{attribute 'linkalways'} 
{attribute 'no_explicit_call' := 'This FB is a CLASS and must be accessed using methods or properties'}
{attribute 'enable_dynamic_creation'}
FUNCTION_BLOCK _ETcVnEdgeDetectionAlgorithm EXTENDS EnumDatatypeBase
VAR
	localData : ETcVnEdgeDetectionAlgorithm;
	activeData : REFERENCE TO ETcVnEdgeDetectionAlgorithm;
	enumBaseDatatype : _DINT(localData);
END_VAR

METHOD PRIVATE AddLocalEnumeration
VAR_INPUT
	Enumeration : T_MAXSTRING;
	Value : ETcVnEdgeDetectionAlgorithm;
END_VAR
AddEnumeration(Enumeration, Value);
END_METHOD

PROPERTY PUBLIC Address : PVOID
GET
Address := ADR(activeData);
END_GET
END_PROPERTY

METHOD PUBLIC ClearReference
VAR_INPUT
END_VAR
activeData REF= localData;
SetBaseDatatypeReference();
END_METHOD

METHOD PUBLIC Clone : I_Datatype
VAR
    pClone : POINTER TO _ETcVnEdgeDetectionAlgorithm;
END_VAR
pClone := __NEW(_ETcVnEdgeDetectionAlgorithm(InitialValue := Value));
Clone := pClone^;
END_METHOD

METHOD FB_init : BOOL
VAR_INPUT
	bInitRetains : BOOL; // if TRUE, the retain variables are initialized (warm start / cold start)
	bInCopyCode : BOOL;  // if TRUE, the instance afterwards gets moved into the copy code (online change)
	InitialValue : ETcVnEdgeDetectionAlgorithm;
END_VAR
localData := InitialValue;
AddBaseDatatype(enumBaseDatatype);
ClearReference();

AddLocalEnumeration('TCVN_EDA_INTERPOLATION', ETcVnEdgeDetectionAlgorithm.TCVN_EDA_INTERPOLATION);
AddLocalEnumeration('TCVN_EDA_APPROX_ERF', ETcVnEdgeDetectionAlgorithm.TCVN_EDA_APPROX_ERF);
AddLocalEnumeration('TCVN_EDA_APPROX_GAUSSIAN', ETcVnEdgeDetectionAlgorithm.TCVN_EDA_APPROX_GAUSSIAN);
END_METHOD

PROPERTY PUBLIC Identifier : T_MAXSTRING
GET
Identifier := 'ETcVnEdgeDetectionAlgorithm';
END_GET
END_PROPERTY

METHOD IsEnumeratorValueEqual : BOOL
VAR_INPUT
	Enumerator : I_KeyValueForwardEnumerator;
END_VAR
VAR
	storedValue : ETcVnEdgeDetectionAlgorithm;
END_VAR
IF NOT Enumerator.TryGet(storedValue) THEN
	RETURN;
END_IF

IsEnumeratorValueEqual := storedValue = activeData;
END_METHOD

METHOD PUBLIC MakeReferenceTo
VAR_INPUT
	ReferenceTarget : REFERENCE TO ETcVnEdgeDetectionAlgorithm;
END_VAR
activeData REF= ReferenceTarget;
SetBaseDatatypeReference();
END_METHOD

METHOD PROTECTED SetBaseDatatypeReference
VAR_INPUT
END_VAR
enumBaseDatatype.MakeReferenceTo(activeData);
END_METHOD

PROPERTY PUBLIC Size : UDINT
GET
Size := SIZEOF(activeData);
END_GET
END_PROPERTY

METHOD TryMakeReferenceTo : BOOL
VAR_INPUT
	Target : I_Datatype;
END_VAR
VAR
	pTargetData : POINTER TO ETcVnEdgeDetectionAlgorithm;
END_VAR
IF NOT IsEquivalentTo(Target) THEN
	RETURN;
END_IF

pTargetData := Target.Address;
activeData REF= pTargetData^;
SetBaseDatatypeReference();
TryMakeReferenceTo := TRUE;
END_METHOD

PROPERTY PUBLIC Value : ETcVnEdgeDetectionAlgorithm
GET
Value := activeData;
END_GET
SET
activeData := Value;
END_SET
END_PROPERTY

END_FUNCTION_BLOCK

(* stored: Version 1.1.0.1, ProductVersion 3.1.4024.13
   POU _ETcVnEdgeDetectionAlgorithm: Id {de3327d9-628b-0db8-070f-b6ec3e9cfed8}, SpecialFunc None
   Folder Core: Id {e035bb8f-f195-0321-2564-328d1d9e6354}
   Folder Protected: Id {24d363fe-2ee2-017f-0644-1bdf48376c97}
   Folder Customize: Id {5e2cb9a4-28a6-0918-2e91-0ebe8bb50e53}
   Folder Constructor: Id {163cf6a0-f511-071e-20fa-813a2df9bf96}
   Folder Private: Id {fa96855c-e46a-09e8-18d9-cd7d699408c7}
   Folder Protected: Id {81f72d85-df5c-0d10-25bf-c5676d71d58f}
   Method AddLocalEnumeration: Id {c7807dc8-fcd2-0167-2c69-db3e14617561}
   Property Address: Id {1c4d0320-6103-0427-3c85-658858caa5d9}
   Get Get: Id {2ceb24b0-bddc-0b13-0661-3c4ac1ff7d2a}
   Method ClearReference: Id {06331ef3-70e5-04b8-06bb-a3e7476cd189}
   Method Clone: Id {93dcc90a-ca49-0669-2de3-8775364a3c48}
   Method FB_init: Id {499c5acc-ee1f-048c-274d-37da243b2af5}
   Property Identifier: Id {73c0b194-9924-0dcf-2ac0-b517abdb4f5b}
   Get Get: Id {2391be6c-42a0-0570-0938-859bb6badf5f}
   Method IsEnumeratorValueEqual: Id {15a04b32-a76a-0a9a-0ce5-ab7589c338e2}
   Method MakeReferenceTo: Id {96185666-00ce-04b4-2ca1-41455ce3c251}
   Method SetBaseDatatypeReference: Id {9d4bfa6b-0ad5-0f35-2704-873b62a7c773}
   Property Size: Id {e13cb641-21be-0973-19f6-6f0b79d34c79}
   Get Get: Id {3bb99596-40a5-0d7a-0259-ebc5370e2b18}
   Method TryMakeReferenceTo: Id {7b1ff354-ecf7-0aaf-01ca-730cbb69bce2}
   Property Value: Id {961ce8f3-bf3e-0537-187a-30ab8e162096}
   Get Get: Id {bb0abdb4-7053-07e8-3dd2-c591c18a5e7c}
   Set Set: Id {08eee3c9-39d1-055b-191e-944ae51f1070} *)
